Staubli VAL3: goSafeHome.pjx

--- goSafeHome.pjx ---
Parameters version=s8.12.1cs9_BS2449 stackSize=200000 millimeterUnit=true
Program file=gosafe.pgx
Program file=start.pgx
Program file=stop.pgx
Data file=goSafeHome.dtx
Library alias=saveData path=Disk://source/saveData/saveData.pjx autoload=true password=
Library alias=rs path=Disk://source/projectSource/robotStatus/robotStatus.pjx autoload=true password=

--- goSafeHome.dtx ---
mdesc mHome = {accel=25, vel=50, decel=25, blend=off}
mdesc mNomSpeed

--- start.pgx ---
program start()
begin
end

--- gosafe.pgx ---
public program gosafe()
  local pointRx l_pHere
  local pointRx l_pHome
  local pointRx l_pMiddle
  local pointRx l_pTrans
  local tool l_tTool
begin
  rs:sTrajStatus="自动回原点过程中"
  setMoveId(1000)
  $jogMode(0)
  link(l_tTool,flange)
  link(l_pTrans,world)
  call saveData:getTool(1,l_tTool)
  l_pHere=here(l_tTool,world)
  l_pHome=jointToPoint(l_tTool,world,saveData:jHome)
  //l_pMiddle=jointToPoint(l_tTool,world,saveData:jMiddle)
  l_pHere.trsf.z=l_pHome.trsf.z


  l_pTrans=l_pHere
  movel(l_pHere,l_tTool,mHome)
  waitEndMove()

  l_pTrans.trsf.x=623
  l_pTrans.trsf.y=0
  l_pTrans.trsf.rx=l_pHere.trsf.rx
  l_pTrans.trsf.ry=l_pHere.trsf.ry
  l_pTrans.trsf.rz=l_pHere.trsf.rz
  movel(l_pTrans,l_tTool,mHome)
  waitEndMove()
  movej(l_pHome,l_tTool,mHome)
  waitEndMove()
  // delay(0)
  rs:sTrajStatus="自动回原点完成,已在待产状态"
end

--- stop.pgx ---
program stop()
begin
end
